// Mitsubishi GX Works2 project: 261012_적산타이머실습   PLC: Q03UDV

PROGRAM MAIN
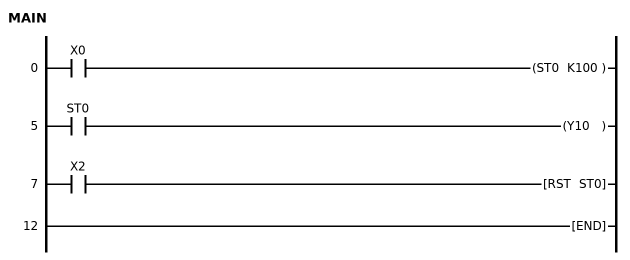
0     LD      X0
      OUT     ST0 K100
5     LD      ST0
      OUT     Y10
7     LD      X2
      RST     ST0
12    END
END_PROGRAM
